Fanuc KAREL source: kc00021.KL

-- PROVISIONAL review KL for V770-1; original PC SHA256 276d2b41bac14e50765a8c684898c1324e88d68160c22b8b678987c8f0521882
-- Incomplete behavior may be omitted. Consult companion uncertainty JSON. Do not deploy.
PROGRAM KC00021
%NOLOCKGROUP
BEGIN
  -- UNRESOLVED_PC offsets 5-18; opcodes 27,27,27,9C,31,23
  -- UNRESOLVED_PC offsets 23-27; opcodes 7F
END KC00021
